Fanuc KAREL source: kb00027.KL

PROGRAM KB00027
%STACKSIZE=65535
%PRIORITY=65535
%NOLOCKGROUP
VAR
P1 : BOOLEAN
P2 : STRING[80]
P3 : INTEGER
BEGIN
P1=TRUE
P2='A'
P3=1
CNC_DYN_DISB(P1,P2,P3)
END KB00027
